// TIA Portal V21 export
// export: Created 2026-11-22T04:06:06.665328Z, ExportSetting WithDefaults, DisplayName Totally Integrated Automation Portal, DisplayVersion V21 Update 3, DisplayName STEP 7 Professional, DisplayVersion V21 Update 3, DisplayName STEP 7 Safety, DisplayVersion V21, DisplayName Tech WebApplication, DisplayVersion V21, DisplayName WinCC Basic/Comfort/Advanced, DisplayVersion V21 Update 3, DisplayName WinCC Unified, DisplayVersion V21 Update 3
ScreenPopup "Popup_C05"  300x200
  ScreenLayer "Layer_0"
    Rectangle "Pop_Back" at 0,0 size 300x200
    TextField "Pop_Title" at 10,10 size 280x20  StyleItem=Text field, Text="Pop-up screen Popup_C05"
    GraphicView "Pop_Graphic" at 10,40 size 120x80  Picture=G_PNG
    IOField "Pop_Value" at 150,60 size 120x30  DataFormat=Decimal, FormatPattern=s99999, Mode=InOutput, StyleItem=I/O field
      ProcessValue := D_Int
    Button "Pop_Close" at 200,160 size 80x22  Mode=Text, StyleItem=Button, TextOff="Close", TextOn="Close"
      on Click: ShowPopupScreen(Name of the screen := , X coordinate := 200, Y coordinate := 120, Display mode := -1, Animation := -1, Animation speed := 1)
